(* IEC 61131-3 sources: SortJet_MasterSPS_Aufbau.fbsproj/11_MMI_Kommunikation/Hegla_Gateway_Komm_FB.fb.st^, 13 files *)

(* ---- CloseSocket.meth.st ---- *)
(* METADATA
{
	"v3Meta": {
		"objectGuid": "9f82718f-b1e3-4bef-8f71-7bc3b9baf787"
	}
}
*)
METHOD CloseSocket : BOOL
//  Closes a socket and sets it invalid.
//  Return: Success of operation
VAR_INPUT
  hSocket: POINTER TO RTS_IEC_HANDLE; // Address of Socket-ID
END_VAR
VAR
  uiResult : UDINT;
END_VAR
CloseSocket := FALSE;
IF ( hSocket <> 0 ) AND ( hSocket^ <> RTS_INVALID_HANDLE )
THEN
  uiResult:= SysSockClose(hSocket^);
  IF uiResult = CmpErrors.Errors.ERR_OK
  THEN
    CloseSocket:= TRUE;
  ELSE
    CloseSocket:= FALSE;
  END_IF
  hSocket^:= RTS_INVALID_HANDLE;
END_IF
END_METHOD

(* ---- Crc32.meth.st ---- *)
(* METADATA
{
	"v3Meta": {
		"objectGuid": "6b6b9ff1-a382-43e7-9f9f-17942cf7a836"
	}
}
*)
METHOD Crc32 : DWORD
VAR_INPUT
  pbpValue : POINTER TO BYTE;
  dwpSize  : DWORD;
END_VAR
VAR
  dwlCrc  : DWORD := 16#FFFFFFFF;
  ilIndex : INT;
END_VAR

// Funktion zur Berechnung einer CRC32-Prüfsumme
dwlCrc := 16#FFFFFFFF;

FOR ilIndex:=1 TO DWORD_TO_INT( dwpSize (*-2*) ) DO
  dwlCrc := SHR(dwlCrc, 8) XOR adwgCrcTable[ ( dwlCrc AND 16#FF ) XOR pbpValue^ ];
  pbpValue := pbpValue + 1;
END_FOR

dwlCrc := dwlCrc XOR 16#FFFFFFFF;

Crc32 := dwlCrc;
END_METHOD

(* ---- GetMessage.act.st ---- *)
(* METADATA
{
	"v3Meta": {
		"objectGuid": "c15a1bbd-8694-42ea-9195-cf52aa2de87e"
	}
}
*)
ACTION GetMessage
IF ( ilAuftraegeAnz = 0 ) THEN
  // CRC32-Summe für die Aufträge prüfen.
  dwAuftragsChecksumme := Crc32( ADR( MmiToSps.smbMessageBlock ), SIZEOF( MmiToSps.smbMessageBlock ) - cSizeOfDWord );
  IF ( HMI_GetDWORD( ADR(MmiToSps.smbMessageBlock.dwCrc32Checksumme)) = dwAuftragsChecksumme ) THEN
    // Nachrichten aus dem Speicher übernehmen und Quitieren
    IF ( ( HMI_GetWORD(ADR(MmiToSps.smbMessageBlock.wCnt2)) <> SpsToMmi.smbMessageBlock.wQuitCnt ) AND
         ( HMI_GetWORD(ADR(MmiToSps.smbMessageBlock.wCnt1)) =  HMI_GetWORD(ADR( MmiToSps.smbMessageBlock.wCnt2 ) ))
       ) THEN
      MemCopy( ADR( asmSpsMessage ), ADR( MmiToSps.smbMessageBlock.asmSpsMessage ), SIZEOF( asmSpsMessage ) );
      ilAuftraegeAnz := WORD_TO_INT(HMI_GetWORD( ADR(MmiToSps.smbMessageBlock.wAnzAuftraege)) );
      IF ilAuftraegeAnz > 5 THEN
        ilAuftraegeAnz := 5; // Schutz vor Array-Überlauf (asmSpsMessage[0..4])
      END_IF
      ilAuftragIndex := 0;
      SpsToMmi.smbMessageBlock.wQuitCnt := HMI_GetWORD(ADR( MmiToSps.smbMessageBlock.wCnt2));
    END_IF;
  END_IF;
END_IF;

// 1 Nachricht pro Zyklus verarbeiten
IF ( ilAuftraegeAnz > 0 ) THEN
  MemCopy( ADR( smlSpsMessage ), ADR( asmSpsMessage[ ilAuftragIndex ] ), SIZEOF( smlSpsMessage ) );
  ilAuftragIndex := ilAuftragIndex + 1;
  // NEU-->
  smlSpsMessage.wAuftrag := HMI_GetWORD(ADR(smlSpsMessage.wAuftrag));
  smlSpsMessage.wLaenge := HMI_GetWORD(ADR(smlSpsMessage.wLaenge));
  // <--NEU
  IF ( MsgInterpret(smlSpsMessage) = FALSE ) THEN
  // smlErrorMsg.wAuftrag   := 32767;
  // smlErrorMsg.wLaenge    := 4;
  // HMI_PutWORD(ADR(smlErrorMsg.awDaten[0]), 3);
  // HMI_PutWORD(ADR(smlErrorMsg.awDaten[1]), smlSpsMessage.wAuftrag);
  // PutMsg( smpSpsMessage := smlErrorMsg, bpTrig := FALSE );

  END_IF
END_IF;
IF ( ilAuftragIndex >= ilAuftraegeAnz ) THEN
  ilAuftraegeAnz := 0;
  ilAuftragIndex := 0;
END_IF;
END_ACTION

(* ---- InMsg.meth.st ---- *)
(* METADATA
{
	"v3Meta": {
		"objectGuid": "cda33201-c5a6-4fe7-8396-38f1974bd209"
	}
}
*)
METHOD InMsg : BOOL
VAR_INPUT
  psmSpsMessage : SpsMessage;
END_VAR
VAR
  i : INT;
  j : INT;
END_VAR

i := smqSpsMessageQueue.iInzeig;
j := (i+1) MOD 25;   // 25 mögliche Queueeinträge möglich

// noch Platz frei ?
IF( j = smqSpsMessageQueue.iOutzeig )THEN
  // Queue ist voll, älteste Nachricht wird verworfen
  smqSpsMessageQueue.iOutzeig := (j+1) MOD 25;
END_IF;

// in jedem Fall eintragen
smqSpsMessageQueue.asmSpsMessage[i] := psmSpsMessage;
smqSpsMessageQueue.iInzeig  := j;

InMsg := TRUE;
END_METHOD

(* ---- M_CloseSocket.meth.st ---- *)
(* METADATA
{
	"v3Meta": {
		"objectGuid": "b05be44e-048d-42d4-abc7-77aa943f133f"
	}
}
*)
METHOD M_CloseSocket : UDINT
VAR_INPUT
END_VAR

CloseSocket(ADR(Client.hSocket));

CloseSocket(ADR(hSocket));
END_METHOD

(* ---- M_ReadMsg_InterpretMsg.meth.st ---- *)
(* METADATA
{
	"v3Meta": {
		"objectGuid": "b9f6b86d-7a91-4709-a115-3d1bc5da6f67"
	}
}
*)
METHOD M_ReadMsg_InterpretMsg : BOOL
VAR_INPUT
END_VAR

M_ReadMsg_InterpretMsg := FALSE;
CASE mhHeader.wType OF

  cMsg_Watchdog:
    // Watchdog Nachricht empfangen
    MmiToSpsMem.wWatchdog := HMI_GetWORD( ADR( bBuffer_Read[4] ) );
    M_ReadMsg_InterpretMsg         := TRUE;

  cMsg_MsgBlock:
    // Messageblock Nachricht empfangen
    // EXC88 keine Buffer Words mehr!
    MemCopy( ADR( MmiToSpsMem.smbMessageBlock.wQuitCnt ),ADR( bBuffer_Read[4] ),cSizeOfWord *3 );

    MemCopy( ADR( MmiToSpsMem.smbMessageBlock.asmSpsMessage[0].wAuftrag ),
             ADR( bBuffer_Read[10] ), SIZEOF( MmiToSpsMem.smbMessageBlock.asmSpsMessage ) ) ;

    // Pointer setzen
    pbCurPos_Read := ADR( bBuffer_Read[10] ) + SIZEOF( MmiToSpsMem.smbMessageBlock.asmSpsMessage );
    MemCopy( ADR( MmiToSpsMem.smbMessageBlock.wCnt2 ), pbCurPos_Read, cSizeOfWord );

    pbCurPos_Read := pbCurPos_Read + 2; // Pointer um 2 Bytes erhöhen
    MemCopy( ADR( MmiToSpsMem.smbMessageBlock.dwCrc32Checksumme ), pbCurPos_Read, cSizeOfDWord );

    M_ReadMsg_InterpretMsg := TRUE;
END_CASE
END_METHOD

(* ---- MsgBegin.act.st ---- *)
(* METADATA
{
	"v3Meta": {
		"objectGuid": "bd949edd-780c-4971-83d6-b01a2ef6b548"
	}
}
*)
ACTION MsgBegin
// Watchdog-Value auf die Struktur übernehmen
Memcopy( ADR( MmiToSps ), ADR( MmiToSpsMem ), cSizeOfWord );

// MessageBlock vom MMI überprüfen
IF( Memcomp( ADR( MmiToSps.smbMessageBlock ), ADR( MmiToSpsMem.smbMessageBlock ), SIZEOF( MmiToSps.smbMessageBlock ) ) <> 0 )THEN
  // Prüfen ob der neue Messageblock vom MMI gültig ist
  dwlChecksumme0 := Crc32( ADR(MmiToSpsMem.smbMessageBlock), SIZEOF( MmiToSps.smbMessageBlock ) - cSizeOfDWord );

  // dwlChecksumme1 :=  MmiToSpsMem.smbMessageBlock.dwCrc32Checksumme;
  dwlChecksumme1 := HMI_GetDWORD( ADR( MmiToSpsMem.smbMessageBlock.dwCrc32Checksumme));

  IF( dwlChecksumme0 = dwlChecksumme1 )THEN
    // neuen MessageBlock vom MMI überbenehmen
    Memcopy( ADR( MmiToSps.smbMessageBlock ), ADR( MmiToSpsMem.smbMessageBlock ), SIZEOF( MmiToSps.smbMessageBlock ));
  END_IF;
END_IF;

Watchdog();
IF( o_b_WatchdogOk )THEN
  GetMessage();
END_IF;
END_ACTION

(* ---- MsgEnd.act.st ---- *)
(* METADATA
{
	"v3Meta": {
		"objectGuid": "0fab3b3e-6742-4984-990c-b65a2821afa3"
	}
}
*)
ACTION MsgEnd
PutMsg( smpSpsMessage := smlSpsMessage_POLL, bpTrig := TRUE );
SendMsg();
IF( Memcomp( ADR( SpsToMmiMem ), ADR( SpsToMmi ), SIZEOF( SpsToMmi ) ) <> 0 )THEN
  Memcopy( ADR( SpsToMmiMem ), ADR( SpsToMmi ), SIZEOF( SpsToMmi ) );
END_IF
IF TCPMain.bpIOAnzeigeAktivieren THEN
  UpdateIoAnzeige();
END_IF
END_ACTION

(* ---- PutMsg.meth.st ---- *)
(* METADATA
{
	"v3Meta": {
		"objectGuid": "e8a694c3-4b92-4b4d-9e51-92b9da22543a"
	}
}
*)
METHOD PutMsg : BOOL
VAR_INPUT
  smpSpsMessage : SpsMessage;
  bpTrig        : BOOL;
END_VAR
VAR
  smlSpsMessage : SpsMessage;
END_VAR

// Nachricht in den Kommunikationspuffer zum MMI eintragen bzw. in die Queue,
//    falls der Kommunikationspuffer belegt ist.

IF( o_b_WatchdogOk <> TRUE )THEN
  RETURN;
END_IF;

// Compilerfehler beim direkten verwenden der Inputvariable bei BLKMOV und MessageIn !?
// Wenn notwenig Drehen, wird in der Funktion GetSpsWord Entscheiden
smlSpsMessage.wAuftrag := HMI_GetWORD(ADR(smpSpsMessage.wAuftrag));
smlSpsMessage.wLaenge  := HMI_GetWORD(ADR(smpSpsMessage.wLaenge));
smlSpsMessage.awDaten  := smpSpsMessage.awDaten; // Die Daten werden in MSGToMMi Aufbereitet

IF( HMI_GetWORD( ADR(MmiToSps.smbMessageBlock.wQuitCnt)) = SpsToMmi.smbMessageBlock.wCnt1 )THEN
  // noch etwas in der Queue ?
  IF( smqSpsMessageQueue.iInzeig <> smqSpsMessageQueue.iOutzeig )THEN
    SpsToMmi.smbMessageBlock.wCnt1 := INT_TO_WORD( WORD_TO_INT( SpsToMmi.smbMessageBlock.wCnt1 ) + 1 );

    // Nachricht 1
    SpsToMmi.smbMessageBlock.wAnzAuftraege := 1;
    Memcopy( ADR( SpsToMmi.smbMessageBlock.asmSpsMessage[0] ), ADR( smqSpsMessageQueue.asmSpsMessage[ smqSpsMessageQueue.iOutzeig ] ), SIZEOF( smlSpsMessage ) );
    smqSpsMessageQueue.iOutzeig := ( smqSpsMessageQueue.iOutzeig + 1 ) MOD 25;

    // Nachricht 2
    IF( smqSpsMessageQueue.iInzeig <> smqSpsMessageQueue.iOutzeig )THEN
      SpsToMmi.smbMessageBlock.wAnzAuftraege := 2;
      Memcopy( ADR( SpsToMmi.smbMessageBlock.asmSpsMessage[1] ), ADR( smqSpsMessageQueue.asmSpsMessage[ smqSpsMessageQueue.iOutzeig ] ), SIZEOF( smlSpsMessage ) );
      smqSpsMessageQueue.iOutzeig := ( smqSpsMessageQueue.iOutzeig + 1 ) MOD 25;
    END_IF;

    // Nachricht 3
    IF( smqSpsMessageQueue.iInzeig <> smqSpsMessageQueue.iOutzeig )THEN
      SpsToMmi.smbMessageBlock.wAnzAuftraege := 3;
      Memcopy( ADR( SpsToMmi.smbMessageBlock.asmSpsMessage[2] ), ADR( smqSpsMessageQueue.asmSpsMessage[ smqSpsMessageQueue.iOutzeig ] ), SIZEOF( smlSpsMessage ) );
      smqSpsMessageQueue.iOutzeig := ( smqSpsMessageQueue.iOutzeig + 1 ) MOD 25;
    END_IF;

    // Nachricht 4
    IF( smqSpsMessageQueue.iInzeig <> smqSpsMessageQueue.iOutzeig )THEN
      SpsToMmi.smbMessageBlock.wAnzAuftraege := 4;
      Memcopy( ADR( SpsToMmi.smbMessageBlock.asmSpsMessage[3] ), ADR( smqSpsMessageQueue.asmSpsMessage[ smqSpsMessageQueue.iOutzeig ] ), SIZEOF( smlSpsMessage ) );
      smqSpsMessageQueue.iOutzeig := ( smqSpsMessageQueue.iOutzeig + 1 ) MOD 25;
    END_IF;

    // Nachricht 5
    IF( smqSpsMessageQueue.iInzeig <> smqSpsMessageQueue.iOutzeig )THEN
      SpsToMmi.smbMessageBlock.wAnzAuftraege := 5;
      Memcopy( ADR( SpsToMmi.smbMessageBlock.asmSpsMessage[4] ), ADR( smqSpsMessageQueue.asmSpsMessage[ smqSpsMessageQueue.iOutzeig ] ), SIZEOF( smlSpsMessage ) );
      smqSpsMessageQueue.iOutzeig := ( smqSpsMessageQueue.iOutzeig + 1 ) MOD 25;
    END_IF;

    SpsToMmi.smbMessageBlock.wCnt2                  := SpsToMmi.smbMessageBlock.wCnt1;
    SpsToMmi.smbMessageBlock.dwCrc32Checksumme      := Crc32( ADR(SpsToMmi.smbMessageBlock ), SIZEOF( SpsToMmi.smbMessageBlock ) - cSizeOfWord );

    IF( NOT bpTrig )THEN
      InMsg( psmSpsMessage:=smlSpsMessage );
    END_IF
  ELSE
    IF( NOT bpTrig )THEN
      InMsg( psmSpsMessage:=smlSpsMessage );
    END_IF;
  END_IF;
ELSE
  IF( NOT bpTrig )THEN
    InMsg( psmSpsMessage:=smlSpsMessage );
  END_IF;
END_IF;
END_METHOD

(* ---- ReadMsg.act.st ---- *)
(* METADATA
{
	"v3Meta": {
		"objectGuid": "f24bca42-101c-4726-904f-63b36c6b8d1a"
	}
}
*)
ACTION ReadMsg
// Receive Data

IF ( bgTcpConnected AND (Client.hSocket <> RTS_INVALID_HANDLE) ) THEN

  //Reset the variables to receive a new MSG
  IF      l_b_ReadMsg_NewMsg
          AND NOT l_b_ReadMsg_Failure
  THEN
    pbCunrrent := ADR( bBuffer_Read[0] );
    l_b_ReadMsg_NewMsg := FALSE;
    l_b_ReadMsg_Body := FALSE;
  END_IF

  //Read the Header Out of the Buffer to get the type of MSG and it's designated length.
  IF  NOT l_b_ReadMsg_NewMsg
      AND NOT l_b_ReadMsg_Body
      AND NOT l_b_ReadMsg_Failure
  THEN
    diLenght  := DWORD_TO_DINT(ADR( bBuffer_Read[0] ) + SIZEOF( mhHeader ) - pbCunrrent);

    diReceived := TcpReceiveData( Client.hSocket, pbCunrrent, diLenght, 0, ADR(tcpLastError) );

    IF ( diReceived >= 0 ) THEN // Daten empfangen
      pbCunrrent := pbCunrrent + LINT_TO_DWORD(diReceived);
    ELSE
      CloseSocket( ADR( Client.hSocket ) );
    END_IF

    diRemaining := DWORD_TO_DINT(ADR( bBuffer_Read[0] ) + SIZEOF( mhHeader) - pbCunrrent);

    IF ( diRemaining = 0 )
    THEN
      // Header Komplett, next step read the body
      mhHeader.wType   := HMI_GetWORD( ADR( bBuffer_Read[0] ) );
      mhHeader.wLenght := HMI_GetWORD( ADR( bBuffer_Read[2] ) );
      IF ( mhHeader.wLenght <= SIZEOF( bBuffer_Read ) - SIZEOF( mhHeader ) ) THEN
        l_b_ReadMsg_Body := TRUE;
      ELSE
        CloseSocket( ADR( Client.hSocket ) );
      END_IF
    ELSIF (diRemaining < 0)
    THEN
      // Fehler in der Datenverabeitung
      CloseSocket( ADR( Client.hSocket ) );
    END_IF
  END_IF

  //After we now how big the body is, we can read it.
  IF      l_b_ReadMsg_Body
          AND NOT l_b_ReadMsg_Failure
  THEN
    diLenght := DWORD_TO_DINT(ADR( bBuffer_Read[SIZEOF(mhHeader)] ) + mhHeader.wLenght - pbCunrrent);

    diReceived := TcpReceiveData( Client.hSocket, pbCunrrent, diLenght, 0, ADR(tcpLastError) );

    IF ( diReceived >= 0 ) THEN // Daten empfangen
      pbCunrrent := pbCunrrent + LINT_TO_DWORD(diReceived);
    ELSE;
      CloseSocket( ADR( Client.hSocket ) );
    END_IF

    diRemaining := DWORD_TO_DINT(ADR( bBuffer_Read[SIZEOF( mhHeader )] ) + mhHeader.wLenght - pbCunrrent);

    IF (diRemaining = 0 ) THEN
      // Daten Komplett
      IF M_ReadMsg_InterpretMsg()
      THEN
        l_b_ReadMsg_NewMsg := TRUE;
      ELSE
        l_b_ReadMsg_NewMsg := TRUE; //Unbekannte Nachricht verwerfen und weiter.
      END_IF;
    ELSIF ( diRemaining < 0 ) THEN
      CloseSocket( ADR( Client.hSocket ) );
    END_IF
  END_IF

ELSE
  //Try to read a new msg, when the connection resets.
  l_b_ReadMsg_NewMsg := TRUE;
  l_b_ReadMsg_Failure := FALSE;
END_IF
END_ACTION

(* ---- SendMsg.act.st ---- *)
(* METADATA
{
	"v3Meta": {
		"objectGuid": "1d0ebe0f-be57-4ced-a649-54fad2d51936"
	}
}
*)
ACTION SendMsg
// --------------------------Datenabgleich wird bei jeder veränderung ausgeführt--------------------------
IF ( bgTcpConnected AND (Client.hSocket <> RTS_INVALID_HANDLE)) THEN

  IF ( MemComp( ADR( SpsToTcp.wWatchdog ), ADR( SpsToMmiMem.wWatchdog ), SIZEOF( SpsToMmiMem.wWatchdog ) ) <> 0 ) THEN
    MemCopy( ADR( SpsToTcp.wWatchdog ), ADR( SpsToMmiMem.wWatchdog ), SIZEOF( SpsToMmiMem.wWatchdog ) );
    bSendWatchDog := TRUE;
  END_IF

  IF ( MemComp( ADR( SpsToTcp.smbMessageBlock ), ADR( SpsToMmiMem.smbMessageBlock ), SIZEOF( SpsToMmiMem.smbMessageBlock ) ) <> 0 ) THEN
    MemCopy( ADR( SpsToTcp.smbMessageBlock ), ADR( SpsToMmiMem.smbMessageBlock ), SIZEOF( SpsToMmiMem.smbMessageBlock ) );
    bSendMsgBlock := TRUE;
  END_IF

  tnSendIoSystem(IN := TRUE,PT := tSendIoSystem);
  IF ( MemComp( ADR( SpsToTcp.ioSystem ), ADR( SpsToMmiMem.ioSystem ), SIZEOF( SpsToMmiMem.ioSystem ) ) <> 0 )
     AND(tnSendIoSystem.Q)
  THEN
    MemCopy( ADR( SpsToTcp.ioSystem ), ADR( SpsToMmiMem.ioSystem ), SIZEOF( SpsToMmiMem.ioSystem ) );
    bSendIoSystem := TRUE;
    tnSendIoSystem(IN := FALSE);
  END_IF

  IF ( MemComp( ADR( SpsToTcp.aucControlSystem ), ADR( SpsToMmiMem.aucControlSystem ), SIZEOF( SpsToMmiMem.aucControlSystem ) ) <> 0 ) THEN
    MemCopy( ADR( SpsToTcp.aucControlSystem ), ADR( SpsToMmiMem.aucControlSystem), SIZEOF( SpsToMmiMem.aucControlSystem ) );
    bSendControlSystem := TRUE;
  END_IF

  IF ( MemComp( ADR( SpsToTcp.aAntrieb ), ADR( SpsToMmiMem.aAntrieb ), SIZEOF( SpsToMmiMem.aAntrieb ) ) <> 0 ) THEN
    MemCopy( ADR( SpsToTcp.aAntrieb ), ADR( SpsToMmiMem.aAntrieb), SIZEOF( SpsToMmiMem.aAntrieb ) );
    bSendDrives := TRUE;
  END_IF
END_IF

IF ( NOT bgTcpConnected ) THEN
  SpsToTcp.wWatchdog := 0;
  SpsToMmi.wWatchdog := 0;
  SpsToMmiMem.wWatchdog := 0;
  MmiToSps.wWatchdog := 0;
  MmiToSpsMem.wWatchdog := 0;
  bTimeOff := FALSE;
  wZyklenOff := 0;
END_IF

// --------------------------Watchdog versenden-------------------------------------------------------
IF bSendWatchDog AND (Client.hSocket <> RTS_INVALID_HANDLE) THEN

  HMI_PutWORD( ADR( mhMsgHeader.wType ), cMsg_Watchdog );
  HMI_PutWORD( ADR( mhMsgHeader.wLenght ), SIZEOF( SpsToTcp.wWatchdog ) );
  HMI_PutWORD( ADR( bBuffer_Send[0] ),SpsToTcp.wWatchdog );

  // Header Versenden
  diSent := TcpSendData( Client.hSocket, ADR( mhMsgHeader ), SIZEOF( mhMsgHeader), ADR(tcpLastError) );
  IF diSent = SIZEOF( mhMsgHeader ) THEN
    // Daten Versenden
    diSent := TcpSendData( Client.hSocket, ADR( bBuffer_Send[0] ), SIZEOF( SpsToTcp.wWatchdog), ADR(tcpLastError) ) ;
    IF diSent = SIZEOF( SpsToTcp.wWatchdog ) THEN
      bSendWatchDog := FALSE;
    ELSIF diSent <> 0 THEN
      IF tcpTrace = 0 THEN
        tcpTrace := 2;
      END_IF
      CloseSocket( ADR( Client.hSocket ) );
    END_IF
  ELSIF diSent <> 0 THEN
    IF tcpTrace = 0 THEN
      tcpTrace := 1;
    END_IF
    CloseSocket( ADR( Client.hSocket ) );
  END_IF
END_IF

// --------------------------MsgBlock versenden-------------------------------------------------------
IF ( bSendMsgBlock AND (Client.hSocket <> RTS_INVALID_HANDLE) ) THEN
  wSendMsgBlock := wSendMsgBlock+1;

  // Daten umkopieren und für die Oberfläche vorbereiten
  // Es kann nicht der gesammte Msg Block 1:1 umkopiert werden weil es bei der Ekelmann Steuerung
  //  nachdem 3 Word und vor dem letzen DWORD des MsgBlock 2 Buffer Bytes gibt

  HMI_PutWORD( ADR( mhMsgHeader.wType ), cMsg_MsgBlock );
  HMI_PutWORD( ADR( mhMsgHeader.wLenght ), 332 );// Original Byte Größe verwenden bei Sizeof() werden BufferBytes mitberechnet

  HMI_PutWORD( ADR( bBuffer_Send[0] ),SpsToTcp.smbMessageBlock.wQuitCnt );
  HMI_PutWORD( ADR( bBuffer_Send[2] ),SpsToTcp.smbMessageBlock.wCnt1 );
  HMI_PutWORD( ADR( bBuffer_Send[4] ),SpsToTcp.smbMessageBlock.wAnzAuftraege );

  MemCopy( ADR( bBuffer_Send[6] ),ADR( SpsToTcp.smbMessageBlock.asmSpsMessage ),SIZEOF( SpsToTcp.smbMessageBlock.asmSpsMessage ) );

  pbCurPos_Send := ADR( bBuffer_Send[6])+ SIZEOF( SpsToTcp.smbMessageBlock.asmSpsMessage );
  HMI_PutWORD( pbCurPos_Send, SpsToTcp.smbMessageBlock.wCnt2 );

  dwCrcTemp :=  Crc32( ADR( bBuffer_Send[0] ), SIZEOF( SpsToTcp.smbMessageBlock ) - cSizeOfWord );

  pbCurPos_Send := pbCurPos_Send +2 ;
  HMI_PutDWORD( pbCurPos_Send,dwCrcTemp );

  // Header versenden
  diSent := TcpSendData( Client.hSocket, ADR( mhMsgHeader ), SIZEOF( mhMsgHeader ), ADR(tcpLastError)  );
  IF diSent = SIZEOF( mhMsgHeader ) THEN
    diSent := TcpSendData( Client.hSocket, ADR( bBuffer_Send[0] ), 332, ADR(tcpLastError)  );
    IF diSent = 332 THEN
      bSendMsgBlock := FALSE;
    ELSIF diSent <> 0 THEN
      IF tcpTrace = 0 THEN tcpTrace := 4; END_IF
      CloseSocket( ADR( Client.hSocket ) );
    END_IF
  ELSIF diSent <> 0 THEN
    IF tcpTrace = 0 THEN tcpTrace := 3; END_IF
    CloseSocket( ADR( Client.hSocket ) );
  END_IF
END_IF

// -------------------------- ConrolSystem versenden-------------------------------------------------------
IF ( bSendControlSystem AND (Client.hSocket <> RTS_INVALID_HANDLE) ) THEN
  wSendControlSystem := wSendControlSystem+1;

  HMI_PutWORD( ADR( mhMsgHeader.wType ), cMsg_ControlSystem );
  HMI_PutWORD( ADR( mhMsgHeader.wLenght ), SIZEOF( SpsToTcp.aucControlSystem ) );

  MemCopy( ADR( bBuffer_Send[0] ), ADR( SpsToTcp.aucControlSystem ), SIZEOF( SpsToTcp.aucControlSystem ) );

  diSent := TcpSendData( Client.hSocket, ADR( mhMsgHeader ), SIZEOF( mhMsgHeader ), ADR(tcpLastError)  );
  // Header Versenden
  IF diSent = SIZEOF( mhMsgHeader ) THEN
    // Daten versenden
    diSent := TcpSendData( Client.hSocket, ADR( bBuffer_Send[0] ), SIZEOF( SpsToTcp.aucControlSystem ), ADR(tcpLastError)  );
    IF diSent = SIZEOF( SpsToTcp.aucControlSystem ) THEN
      bSendControlSystem := FALSE;
    ELSIF diSent <> 0 THEN
      IF tcpTrace = 0 THEN tcpTrace := 6; END_IF
      CloseSocket( ADR( Client.hSocket ) );
    END_IF
  ELSIF diSent <> 0 THEN
    IF tcpTrace = 0 THEN tcpTrace := 5; END_IF
    CloseSocket( ADR( Client.hSocket ) );
  END_IF
END_IF

// -------------------------- IO's versenden-------------------------------------------------------

IF ( bSendIoSystem AND (Client.hSocket <> RTS_INVALID_HANDLE) ) THEN
  wSendIoSystem := wSendIoSystem+1;

  HMI_PutWORD( ADR( mhMsgHeader.wType ), cMsg_IOSystem );
  HMI_PutWORD( ADR( mhMsgHeader.wLenght ), SIZEOF( SpsToTcp.ioSystem ) );

  MemCopy( ADR( bBuffer_Send[0] ), ADR( SpsToTcp.ioSystem ), SIZEOF( SpsToTcp.ioSystem ) );

  // Header versenden
  diSent := TcpSendData( Client.hSocket, ADR( mhMsgHeader ), SIZEOF( mhMsgHeader ), ADR(tcpLastError) );
  IF diSent = SIZEOF( mhMsgHeader ) THEN
    // Daten Versenden
    diSent := TcpSendData( Client.hSocket, ADR( bBuffer_Send[0] ), SIZEOF( SpsToTcp.ioSystem ), ADR(tcpLastError) );
    IF diSent = SIZEOF( SpsToTcp.ioSystem ) THEN
      bSendIoSystem := FALSE;
    ELSIF diSent <> 0 THEN
      IF tcpTrace = 0 THEN tcpTrace := 66; END_IF
      CloseSocket( ADR( Client.hSocket ) );
    END_IF
  ELSIF diSent <> 0 THEN
    IF tcpTrace = 0 THEN tcpTrace := 55; END_IF
    CloseSocket(ADR(Client.hSocket));
  END_IF
END_IF

IF ( FALSE AND  bSendDrives AND (Client.hSocket <> RTS_INVALID_HANDLE) ) THEN

  HMI_PutWORD( ADR( mhMsgHeader.wType ), cMsg_Drives );
  HMI_PutWORD( ADR( mhMsgHeader.wLenght ), SIZEOF( SpsToTcp.aAntrieb ) );

  pbCurPos_Send := ADR( bBuffer_Send[0] );

  FOR i := 0 TO 18 BY 1 DO

    FOR j := 0 TO 8 BY 1 DO

      HMI_PutWORD( pbCurPos_Send,SpsToTcp.aAntrieb[i].awPAE[j] );
      pbCurPos_Send := pbCurPos_Send +2;
      HMI_PutWORD( pbCurPos_Send,SpsToTcp.aAntrieb[i].awPAA[j] );
      pbCurPos_Send := pbCurPos_Send +2;
    END_FOR;

  END_FOR;

  // Header Versenden
  diSent := TcpSendData( Client.hSocket, ADR( mhMsgHeader ), SIZEOF( mhMsgHeader ), ADR(tcpLastError) );
  IF diSent = SIZEOF( mhMsgHeader ) THEN
    // Daten Versenden
    diSent := TcpSendData( Client.hSocket, ADR( bBuffer_Send[0] ), SIZEOF( SpsToTcp.aAntrieb ), ADR(tcpLastError) );
    IF diSent = SIZEOF( SpsToTcp.aAntrieb ) THEN
      bSendDrives := FALSE;
    ELSIF diSent <> 0 THEN
      CloseSocket(ADR(Client.hSocket));
    END_IF
  ELSIF diSent <> 0 THEN
    CloseSocket(ADR(Client.hSocket));
  END_IF
END_IF
END_ACTION

(* ---- TCP_Server.act.st ---- *)
(* METADATA
{
	"v3Meta": {
		"objectGuid": "305dcaac-e980-4088-8579-24e649819553"
	}
}
*)
ACTION TCP_Server
IF bInit THEN

  IF ( hSocket <> RTS_INVALID_HANDLE ) THEN
    IF ( Client.hSocket <> RTS_INVALID_HANDLE ) THEN
      CloseSocket( ADR(Client.hSocket) );
      Client.stIPAddress := '';
    END_IF

    CloseSocket( ADR(hSocket) );
  END_IF

  bgTcpConnected := FALSE;
  tonlOpenForClient(IN := FALSE);
  bInit := FALSE;
ELSE
  tonlOpenForClient(IN := TRUE,PT := T#5000MS);

  // Server Socket öffnen
  IF  hSocket = RTS_INVALID_HANDLE
      AND tonlOpenForClient.Q
  THEN
    hSocket := TcpServerOpenSocket(4444, 1);
  ELSIF tonlOpenForClient.Q THEN
    // Auf Client verbindung warten
    IF Client.hSocket = RTS_INVALID_HANDLE
    THEN
      bgTcpConnected := FALSE;
      Client := TcpServerWaitForConnect(hSocket, 0);
    ELSE
      bgTcpConnected := TRUE;
    END_IF;

  END_IF
END_IF

blVerbindungReset :=
                    (NOT o_b_WatchdogOk) AND
                    (wZyklenOff > 30) AND
                    (Client.hSocket <> RTS_INVALID_HANDLE) AND
                    (NOT tnlVerbindungReset.Q);

tnlVerbindungReset(IN := blVerbindungReset, PT := WORD_TO_TIME(wlVerbindungReset));
rtlVerbindungReset(CLK := tnlVerbindungReset.Q);

IF (rtlVerbindungReset.Q) THEN
  // SendMsg.berror := FALSE;
  CloseSocket(ADR(Client.hSocket));
  Client.stIPAddress := '';
END_IF;

ReadMsg();
END_ACTION

(* ---- WatchDog.act.st ---- *)
(* METADATA
{
	"v3Meta": {
		"objectGuid": "4a5dc8cc-233c-4d19-b434-5bbaf5270e22"
	}
}
*)
ACTION WatchDog
ilDiff := WORD_TO_INT( MmiToSps.wWatchdog ) - WORD_TO_INT( SpsToMmi.wWatchdog );
tlTimeDiff := TIME() - tlTimeOut;

IF (tlTimeDiff > T#5s) THEN
  bTimeOff := TRUE;
  wZyklenOff := wZyklenOff + 1;
  IF ( ilDiff <> 1 ) THEN
    wlWatchdogOk := wlWatchdogOk + 1;
  END_IF
END_IF

IF ( ilDiff <> 1 ) THEN

  IF ( tlTimeDiff > T#5s ) THEN
    // Kommunikationstimeout erreicht
    IF (wZyklenOff>30)
    THEN
      o_b_WatchdogOk := FALSE;
    END_IF
  END_IF

ELSE

  IF ( NOT o_b_WatchdogOk ) THEN
    dwlCrc32Value        := Crc32(ADR( MmiToSps.smbMessageBlock ), SIZEOF( MmiToSps.smbMessageBlock ) - cSizeOfDWord );
    dwAuftragsChecksumme_WatchDog := HMI_GetDWORD(ADR(MmiToSps.smbMessageBlock.dwCrc32Checksumme));
    IF ( ( dwlCrc32Value = dwAuftragsChecksumme_WatchDog ) AND
         ( MmiToSps.smbMessageBlock.wCnt1 = HMI_GetWORD(ADR(SpsToMmi.smbMessageBlock.wQuitCnt))) AND
         ( MmiToSps.smbMessageBlock.wCnt2 = HMI_GetWORD(ADR(SpsToMmi.smbMessageBlock.wQuitCnt))) AND
         ( MmiToSps.smbMessageBlock.wQuitCnt = HMI_GetWORD(ADR(SpsToMmi.smbMessageBlock.wCnt1))) AND
         ( MmiToSps.smbMessageBlock.wQuitCnt = HMI_GetWORD(ADR(SpsToMmi.smbMessageBlock.wCnt2)))
       ) THEN
      o_b_WatchdogOk := TRUE;
      wZyklenOff     := 0;
      bTimeOff       := FALSE;
    END_IF
  END_IF

  tlTimeOut := TIME();

END_IF
IF ( NOT o_b_WatchdogOk ) THEN
  SpsToMmi.smbMessageBlock.wCnt1    := SpsToMmi.smbMessageBlock.wCnt2;
  SpsToMmi.smbMessageBlock.wQuitCnt := HMI_GetWORD(ADR(MmiToSps.smbMessageBlock.wCnt2));

  SpsToMmi.smbMessageBlock.dwCrc32Checksumme := Crc32( ADR( SpsToMmi.smbMessageBlock ), SIZEOF( SpsToMmi.smbMessageBlock ) - cSizeOfDWord );

END_IF
SpsToMmi.wWatchdog := MmiToSps.wWatchdog;
END_ACTION
